(* IEC 61131-3 sources: SRCI_CLIENT_PLC/RobotLibrary/Library/POUs/Read/MC_ReadActualPositionCyclic/Structures, 2 files *)

(* ---- ReadActualPositionCyclicOutCmd.st ---- *)
{attribute 'pack_mode' := '1'}
// -------------------------------------------------------------------------
//  SRCI Robot Library
// -------------------------------------------------------------------------
//
//  Object:      ReadActualPositionCyclicOutCmd
//  Author:      Thorsten Brach
//  Date:        2024-08-09
//
//  Description:
//
//
//  Copyright:
//    (C) 2024 Thorsten Brach. All rights reserved
//             Licensed under the MIT License.
//
//  Disclaimer:
//    This project is provided without any guarantee and can be used for
//    private and commercial purposes. Any use is at the user’s
//    own risk and responsibility.
//
// -------------------------------------------------------------------------
TYPE ReadActualPositionCyclicOutCmd :
STRUCT
  /// TRUE, while the output CartesianPosition returns valid values
  ReadingCartesianPosition    : BOOL;
  /// TRUE, while the output ExtCartesianPosition returns valid values
  ReadingCartesianPositionExt : BOOL;
  /// TRUE, while the output JointPosition returns valid values
  ReadingJointPosition        : BOOL;
  /// TRUE, while the output ExtJointPosition returns valid values
  ReadingJointPositionExt     : BOOL;
  /// Tool and frame index of currently used tool and frame according to Table 6-40
  CurrentCoordinateSystem     : CoordinateSystem;
  /// Cyclically returned, absolute coordinates of current position in selected coordinate systems (see input parameters ToolNo and FrameNo)
  CartesianPosition           : RobotCartesianPosition;
  /// Cyclically returned, absolute coordinates of current position in selected coordinate systems (see input parameters ToolNo and FrameNo)
  CartesianPositionShort      : RobotCartesianPositionShort;
  /// Cyclically returned, absolute cartesian position of the external axes of the robot
  CartesianPositionExt        : RobotCartesianPositionExt;
  /// Tool and frame index of returned position according to Table 6-40
  CoordinateSystem            : CoordinateSystem;
  /// Cyclically returned, absolute joint position of the robot in Joint position
  JointPosition               : RobotJointPosition;
  /// Cyclically returned, absolute short joint position of the robot in Joint position
  JointPositionShort          : RobotJointPositionShort;
  /// Cyclically returned, absolute extended joint position of the external axes of the robot
  JointPositionExt            : RobotJointPositionExt;
END_STRUCT
END_TYPE

(* ---- ReadActualPositionCyclicParCmd.st ---- *)
{attribute 'pack_mode' := '1'}
// -------------------------------------------------------------------------
//  SRCI Robot Library
// -------------------------------------------------------------------------
//
//  Object:      ReadActualPositionCyclicParCmd
//  Author:      Thorsten Brach
//  Date:        2024-08-09
//
//  Description:
//
//
//  Copyright:
//    (C) 2024 Thorsten Brach. All rights reserved
//             Licensed under the MIT License.
//
//  Disclaimer:
//    This project is provided without any guarantee and can be used for
//    private and commercial purposes. Any use is at the user’s
//    own risk and responsibility.
//
// -------------------------------------------------------------------------
TYPE ReadActualPositionCyclicParCmd :
STRUCT
  /// Set TRUE (default) to activate cyclic transmission of cartesian position without external axes
  ReadCartesianPosition       : BOOL := TRUE; // ST-FIX F156: spec 6.1.6 table 6-41: TRUE (default)
  /// Set TRUE to activate cyclic transmission of external axes values of cartesian position -  Default: False
  ReadCartesianPositionExt    : BOOL;
  ///Index of tool of returned position
  /// •     -1: Currently used tool on RC
  /// •      0: Flange (default)
  /// • 1..254: Tool frames
  ToolNo                      : INT;
  /// Index of frame of returned position
  /// •     -1: Currently used frame on RC
  /// •      0: WCS (default)
  /// • 1..254: User frames
  FrameNo                     : INT;
  /// Set TRUE (default) to activate cyclic transmission of joint position without external axes
  ReadJointPosition           : BOOL := TRUE; // ST-FIX F156: spec 6.1.6 table 6-41: TRUE (default)
  /// Set TRUE to activate cyclic transmission of external axes values of joint position - Default: False
  ReadJointPositionExt        : BOOL;
END_STRUCT
END_TYPE
